Fanuc KAREL source: kt00580.KL

-- PROVISIONAL review KL for V940-1; original PC SHA256 7c07110a25a996b513aed10d9267011bc0d2737f9e634bb99979cada242fc78f
-- Incomplete behavior may be omitted. Consult companion uncertainty JSON. Do not deploy.
PROGRAM KT00580
%NOLOCKGROUP
VAR
  I2 : INTEGER
-- UNRESOLVED_DECL V1 type=000013
-- UNRESOLVED_DECL OUT type=000013
BEGIN
  -- V9_ZERO_TABLE_METADATA_HINT layout=0001; no indexed target words; source/name/runtime held
  -- UNRESOLVED_PC offsets 5-20; opcodes 2E,22,32,35
  -- UNRESOLVED_PC offsets 25-36; opcodes 2E,23
  -- UNRESOLVED_PC offsets 41-63; opcodes 49,21,8D,4A
  -- UNRESOLVED_PC offsets 68-72; opcodes 7F
END KT00580
